// TIA Portal V21 export
// export: Created 2026-10-23T20:42:28.3927301Z, ExportSetting WithDefaults, DisplayName Totally Integrated Automation Portal, DisplayVersion V21 Update 1, DisplayName SINAMICS Startdrive Advanced, DisplayVersion V21 HF2, DisplayName SINAMICS Startdrive G110M, G120, G120C, G120D, G120P, G115D, DisplayVersion V21 HF2, DisplayName SINAMICS Startdrive G130, G150, S120, S150, G200, G220, S200, S210, S220, Innomotics MVD, DisplayVersion V21 HF2, DisplayName STEP 7 Professional, DisplayVersion V21 Update 1, DisplayName STEP 7 Safety, DisplayVersion V21, DisplayName Tech WebApplication, DisplayVersion V21, DisplayName WinCC Basic/Comfort/Advanced, DisplayVersion V21 Update 1, DisplayName WinCC Unified, DisplayVersion V21 Update 1
FUNCTION "FC_SclAtOverlay" : Byte   // FC3, SCL
TITLE = AT overlay in a standard block
{ S7_Optimized_Access := 'FALSE' }
VERSION : 0.1
// AT overlays are only allowed in blocks without optimized access
// stored: AutoNumber true, IsIECCheckEnabled false, SetENOAutomatically false, UDAEnableTagReadback false
   VAR_INPUT
      InWord : Word;   // Word to split into bytes
   END_VAR
   VAR_OUTPUT
      HighByte : Byte;   // High byte of InWord
   END_VAR
   VAR_TEMP
      RawWord : Word;   // Raw word
      RawBytes AT RawWord : Array[0..1] of Byte;   // Overlay of RawWord as bytes
   END_VAR
BEGIN

       REGION AT overlay
           #RawWord := #InWord;
           #HighByte := #RawBytes[0];
           #FC_SclAtOverlay := #RawBytes[1];
       END_REGION
END_FUNCTION
